TYPE stAI_DataPoint_APP :
STRUCT
	bActivateLimitCheck			: BOOL;
	bActivateValueChangeCheck	: BOOL;
	fAppValue			: REAL;
	fAppMinValue		: REAL;
	fAppMaxValue		: REAL;
	fAppValueChangeDelta: REAL; 
	tChangeDeltaTime	: TIME;
END_STRUCT
END_TYPE

(* stored: Version 1.1.0.1
   DUT stAI_DataPoint_APP: Id {809b3e21-c3ac-4ad4-9e80-e671e306cd7e} *)
